(*
SPDX-FileCopyrightText: © 2026 Oleksandr Tiutyk <trofimich@gmail.com>
SPDX-License-Identifier: MIT
License: https://opensource.org/license/mit
*)

(*!
<summary>Creates dynamic custom workflow instances and embedded dependencies.</summary>
<description>
Creation transfers exclusive ownership of a fresh unshared instance to the caller.
Return zero for an unknown type name.
</description>
*)
INTERFACE IWorkflowDependencyFactory

(*!
<summary>Creates a fresh unowned dynamic custom workflow or embedded dependency.</summary>
<description>Return zero for an unknown type name.</description>
<param name="typeName">Qualified PLC type name.</param>
*)
METHOD CreateDependency : TOF_Core.IObject
VAR_INPUT
	typeName : STRING(255);
END_VAR
END_METHOD

END_INTERFACE

(* stored: Version 1.1.0.1
   Itf IWorkflowDependencyFactory: Id {e8f1b78d-8986-4cd6-ac40-f4a35ba7982b}
   Method CreateDependency: Id {7d208a81-b0a8-4b8b-b8af-30ed6a6cfcdb} *)
